// Erreur rendue par le chargeur (docs/05 § 10)
{attribute 'pack_mode' := '1'}
TYPE ST_DeployError :
STRUCT
    nCode : UINT;                   // voir FB_Loader
    nStation : USINT;               // 0 = machine
    nTable : USINT;
    nInstr : INT;
    nObject : UINT;
    nDetail : UDINT;
END_STRUCT
END_TYPE

(* stored: Version 1.1.0.1, ProductVersion 3.1.4024.12
   DUT ST_DeployError: Id {5df01c2f-5556-50ea-b436-e27867f48a5b} *)
